(* IEC 61131-3 sources: SortJet_MasterSPS_Aufbau.fbsproj/02_Global Variables, 6 files *)

(* ---- Global_Vars.gvl ---- *)
(* METADATA
{
	"v3Meta": {
		"objectGuid": "27064ae7-2a3c-4a30-8168-a3ab5c131298"
	}
}
*)
{attribute 'allow_unqualified_access'}
NAMESPACE Global_Vars
// Vor StationBasisParameter (Slot 310) initialisieren, dort werden bgFALSE/rgNULL verwendet
{attribute 'global_init_slot' := '295'}
VAR_GLOBAL
//-------------------------------------------------------------------------------------------------
// ALLGEMEINE VARIABLEN
//-------------------------------------------------------------------------------------------------

  // Pointer auf alle Antriebe
  pgAntriebe   : ARRAY[0..65] OF Rexroth_ctrlX_Drive_Eckelmann_MC_V01_02_02;
  bgEtherCatOK : BOOL;

  // Aktivieren \ Deaktivieren des SystemChecks
  bgSystemCheck : ARRAY[cERSTER_AUTOMATIKKREIS..cLETZTER_AUTOMATIKKREIS] OF BOOL := [ cANZAHL_AUTOMATIKKREISE(TRUE) ]; // SystemCheck [AutomatikKreis 1]: FALSE -> Der SystemCheck wird sofort quittiert  TRUE -> SystemCheck wird normal ausgefuehrt

  // Prüfung ob Reset in einem AK aktiv ist
  agbResetAktiv : ARRAY [cERSTER_AUTOMATIKKREIS..cLETZTER_AUTOMATIKKREIS] OF BOOL;

  bgSimulationSiKreisGeschlossen : ARRAY[cERSTER_SICHERHEITSKREIS..cLETZTER_SICHERHEITSKREIS] OF BOOL; // Damit synchronisiert wird, müssen die SKs geschlossen sein - da dies manchmal nicht gegeben ist, kann hiermit

  bgMeldungStromschienenUeberbrueckung : BOOL := FALSE;

  wgStatusPuffer101Oben    : WORD;
  wgStatusPuffer102Unten   : WORD;
  wgStatusPuffer103Oben    : WORD;
  wgStatusPuffer104Unten   : WORD;
  wgStatusTorOben          : WORD;
  wgStatusTorUnten         : WORD;
  // Override für ALLE Achsen - 100 = 100% ; 50 = 50% ;
  rgMaschinenGeschwindigkeitsOverride : REAL := 100;

  (* Hinweis:
     - Pointer- Konstanten [Muessen Global definiert werden]
       => Nicht veraendern
  *)
  bgShuttleEintransportSperren             : ARRAY[cERSTES_SHUTTLE..cLETZTES_SHUTTLE] OF BOOL;
  bgShuttleAustransportSperren             : ARRAY[cERSTES_SHUTTLE..cLETZTES_SHUTTLE] OF BOOL;

  (* Hinweis:
     - Pointer- Konstanten [Muessen Global definiert werden]
       => Nicht veraendern
  *)
  bgTRUE      : BOOL  := TRUE;
  bgFALSE     : BOOL  := FALSE;
  rgNULL      : REAL  := 0;
  wgNULL      : WORD  := 0;

  (* Hinweis:
     - Das Log-Level bestimmt ob und wie die Fehlermeldung geworfen werden->
       Level 0 :=  Nur die übergeordneteten Bausteine werfen einen Fehler
       Level 1 :=  Übergeordnetete Bausteine + Station werfen einen Fehler
       Level 2 :=  Übergeordnetete Bausteine + Station + Unterbausteine werfen einen Fehler
  *)
  wgLogLevel : WORD := 0;
  bgTSLog    : BOOL := TRUE;

  bgStepLogging : BOOL := FALSE;

  Visu_Start_Auto          : BOOL;
  Visu_Notaus_OK           : BOOL := FALSE;

  // Globale Einstellungen
  bgInitialisierungUeberbruecken           : BOOL := FALSE; // Init überspringen
  bgInbetriebnahmeBit                      : BOOL := FALSE; // Inbetriebnahme de/aktivieren
  bgHornAktivieren                         : BOOL := FALSE;  // Horn / Hupe an der Anlage de/aktivieren
  bgSicherheitstechnikBruecken             : BOOL := FALSE; // Inbetriebnahme de/aktivieren
  bgMMIBruecken                            : BOOL := FALSE;
  bgDeaktiviereWatchIOs                    : BOOL := FALSE;
  bgSPS_SIMULATION                         : BOOL := FALSE;
  rgSimScheibenlaenge                      : REAL := 1000.0; // Simulation (bgSPS_SIMULATION): virtuelle Scheibenlaenge [mm] fuer Scheibenmessung und Restwegmessung der simulierten Antriebe
  bgTransfershuttleVortransportAktivieren  : BOOL := FALSE;  // Quittierung des Vortransportauftrags (Ohne Ablauf)
  bgNotHalt_SPS_OK                         : BOOL := TRUE;

  // Ausgaenger - Blink -
  gbFlashbit02sec  : BOOL;
  gbFlashbit05sec  : BOOL;
  gbFlashbit1sec   : BOOL;
  gbFlashbit03sec  : BOOL;
  gbFlashbit12sec  : BOOL;

  // Verfahrueberwachung
  abgVerfahrfreigabeShuttle                    : ARRAY[cERSTES_SHUTTLE..cLETZTES_TRANSFERSHUTTLE] OF BOOL;

  // Init
  M_Init_Ok        : BOOL;

  // Automatikkreise [Speicher - Shuttle - Transfershuttle - ggf. Perepherie
  M_Automatik_Aktiv                         : ARRAY[cERSTER_AUTOMATIKKREIS..cLETZTER_AUTOMATIKKREIS] OF BOOL;
  tonAutomatik_Aktiv                        : ARRAY[cERSTER_AUTOMATIKKREIS..cLETZTER_AUTOMATIKKREIS] OF TON;

  // SystemCheck:
  //   - neue Strukturen aufrufen
  abgDateStationCheck  : ARRAY[101..cLETZTE_STATION, cWAND_1..cANZAHL_WAENDE] OF Auftragsdaten_ST; // Daten die fuer den SystemCheck gebraucht werden

//-------------------------------------------------------------------------------------------------
// ALLGEMEINE STRUKTUREN
//-------------------------------------------------------------------------------------------------
  igIndexFaecherwagenDatenEmpfangen : INT := 0;
  igIndexFaecherwagenDatenSenden    : INT := 0;

  (* Hinweis:
     - Puffer in der Shuttlebahn
  *)
  wgStatusPuffer                       : ARRAY[cERSTES_SHUTTLE..cLETZTES_SHUTTLE] OF WORD;

  (* Hinweis:
     - Allgemeine Konstanten aus der Mathematik
  *)
// *************************************************************************************************
  (* Hinweis:
     - Allgemeine Konstanten aus der Mathematik
  *)
  Mathe : CONSTANTS_MATH;

//-------------------------------------------------------------------------------------------------
// HANDFUNKTIONEN
//-------------------------------------------------------------------------------------------------

  // STATION
  adwgHandfunktionenStationen             : ARRAY[cERSTE_STATION..cLETZTE_STATION] OF DWORD;

  // SHUTTLE
  adwgHandfunktionenShuttle               : ARRAY[cERSTES_SHUTTLE..cLETZTES_SHUTTLE] OF DWORD;

  // TRANSFERSHUTTLE
  adwgHandfunktionenTransfershuttle       : ARRAY[cERSTES_TRANSFERSHUTTLE..cLETZTES_TRANSFERSHUTTLE] OF DWORD;

  // FAECHERWAGENSTATION
  adwgHandfunktionenFaecherwagenStationen : ARRAY[cERSTE_FAECHERWAGENSTATIONS_NR..cLETZTE_FAECHERWAGENSTATIONS_NR] OF DWORD;

//-------------------------------------------------------------------------------------------------
// SYSTEMCHECK
//-------------------------------------------------------------------------------------------------
  wgAnzahlSystemcheckZyklen              : WORD; //  Wird automatisch erkannt

END_VAR
END_NAMESPACE

(* ---- Konstanten.gvl ---- *)
(* METADATA
{
	"v3Meta": {
		"objectGuid": "aefcf88b-f8e6-4fd5-9d29-077a37aead0e"
	}
}
*)
{attribute 'allow_unqualified_access'}
NAMESPACE Konstanten
VAR_GLOBAL CONSTANT

  // Konstanten für die Profibus Master (falls mehrere vorhanden sind)
  cPROFIBUSMASTER_1 : BYTE := 0;
  cPROFIBUSMASTER_2 : BYTE := 1;

  // Konstanten als Ersatz für sizeof
  cSizeOfByte  : WORD := 1;
  cSizeOfWord  : WORD := 2;
  cSizeOfDWord : WORD := 4;
  cSizeOfSInt  : WORD := 1;
  cSizeOfUSInt : WORD := 1;
  cSizeOfInt   : WORD := 2;
  cSizeOfUInt  : WORD := 2;
  cSizeOfDInt  : WORD := 4;
  cSizeOfUDInt : WORD := 4;
  cSizeOfReal  : WORD := 0;

  cMillisecToSec    : WORD  := 1000;
  cMillisecToMinute : WORD  := 60000;

//-------------------------------------------------------------------------------------------------
// SYSTEMCHECK
//-------------------------------------------------------------------------------------------------
  cMAX_ANZAHL_SYSTEMCHECKZYKLEN : WORD := 6;

  // Maximale Anzahl konfigurierbarer Ueberwachungsquellen fuer bpShuttleAnhalten pro Shuttle
  cMAX_SHUTTLE_ANHALTEN_QUELLEN  : WORD := 6;

//-------------------------------------------------------------------------------------------------
// BIT- MASKEN
//-------------------------------------------------------------------------------------------------

  (* Hinweis:
     - Bit Maske
  *)
  // 5432109876543210 ---
  Maske_Bit_0  : WORD := 2#0000000000000001 ;
  Maske_Bit_1  : WORD := 2#0000000000000010 ;
  Maske_Bit_2  : WORD := 2#0000000000000100 ;
  Maske_Bit_3  : WORD := 2#0000000000001000 ;
  Maske_Bit_4  : WORD := 2#0000000000010000 ;
  Maske_Bit_5  : WORD := 2#0000000000100000 ;
  Maske_Bit_6  : WORD := 2#0000000001000000 ;
  Maske_Bit_7  : WORD := 2#0000000010000000 ;
  Maske_Bit_8  : WORD := 2#0000000100000000 ;
  Maske_Bit_9  : WORD := 2#0000001000000000 ;
  Maske_Bit_10 : WORD := 2#0000010000000000 ;
  Maske_Bit_11 : WORD := 2#0000100000000000 ;
  Maske_Bit_12 : WORD := 2#0001000000000000 ;
  Maske_Bit_13 : WORD := 2#0010000000000000 ;
  Maske_Bit_14 : WORD := 2#0100000000000000 ;
  Maske_Bit_15 : WORD := 2#1000000000000000 ;

  // ### KONFIGURIEREN ###

  (* Hinweis:
     - Die folgende Constante darf nicht vergrößert werden, weil es sonst zu einem
       Ueberlauf in der Nachrichtenstruktur kommt
  *)
  cMaxScheibenBeiScheibenMessung  : WORD := 10;

  cMELDUNGScheibe                 : WORD := 0;
  cMAXSCHEIBE                     : WORD := 4;
  cDEFAULTSCHEIBE                 : WORD := 5;
  cMODELLSCHEIBE                  : WORD := 6;

  cGLASDICKEBIS16MM               : WORD := 10;
  cGLASDICKEBIS23MM               : WORD := 11;
  cGLASDICKEBIS29MM               : WORD := 12;

  GLASSTAERKE_DEFAULT_MIN         : WORD := WORD#3;
  GLASSTAERKE_DEFAULT_MAX         : WORD := WORD#14;

  // FAECHERWAGENSTATION
  cEINSCHLEUSESTATION : WORD := 1;
  cPUFFERSTATION      : WORD := 2;
  cFUELLSTATION       : WORD := 3;
  cAUSSCHLEUSESTATION : WORD := 4;
  cKIPPSTATION        : WORD := 5;
  cHUBSTATION         : WORD := 6;
  cENTNAHMESTATION: BOOL := TRUE;

  (* Hinweis:
     - Konstanten fuer das Drehkreuz
  *)
  cGLASDEFAULT : WORD := 0;
  cGLASDREHEN  : WORD := 1;

  (* Hinweis:
     - Grad-Konstanten fuer das Drehkreuz
  *)
  cPOSITION_0Grad    : WORD := 0;
  cPOSITION_90Grad   : WORD := 90;
  cPOSITION_180Grad  : WORD := 180;
  cPOSITION_270Grad  : WORD := 270;
  cPOSITION_360Grad  : WORD := 360;
  rgPOSITION_0Grad   : REAL := REAL#0;
  rgPOSITION_90Grad  : REAL := REAL#90;
  rgPOSITION_180Grad : REAL := REAL#180;
  rgPOSITION_270Grad : REAL := REAL#270;
  rgPOSITION_360Grad : REAL := REAL#360;

  (* Hinweis:
     - Modus wie der FB den Antrieb ansteuern soll
  *)
  cMODUS_MASTER_SLAVE : BYTE := 0;
  cMODUS_HAND         : BYTE := 1;
  cMODUS_RESTWEG      : BYTE := 2;

  (* Hinweis:
     - Unterscheidung Speicher-Einlaufbereich und Speicher-Auslaufbereich
  *)
  cSPEICHER_EINLAUFSEITE : BYTE := 1;
  cSPEICHER_AUSLAUFSEITE : BYTE := 2;

  // Zuweisungskonstanten
  cNULL              : WORD := 0;
  cNULL_WORD_ARRAY   : ARRAY [0..3] OF WORD  :=[ 4(0)];
  cNULL_DWORD_ARRAY  : ARRAY [0..3] OF DWORD :=[ 4(0)];

  cFUEHRUNGSWAGEN    : WORD := 1;
  cZAHNSTANGE        : WORD := 2;

  cSCHMIERKREIS_1    : WORD := 1;
  cSCHMIERKREIS_2    : WORD := 2;
  cSCHMIERKREIS_1_2  : WORD := 3;

//-------------------------------------------------------------------------------------------------
// FOLGEAUFTRAGSTYPEN
//-------------------------------------------------------------------------------------------------
  cFOLGEAUFTRAG_NICHT_AKTIV : WORD := 0;
  cFOLGEAUFTRAG_AKTIV       : WORD := 1;

//-------------------------------------------------------------------------------------------------
// S T A R T - Beladungs- Typ fuer die Shuttle / Stationen nach einem SystemCheck
//-------------------------------------------------------------------------------------------------
  cSTATUS_STATION_FREI              : WORD := 0;
  cSTATUS_STATION_BELEGT            : WORD := 1;
  cSTATUS_STATION_BELEGT_NACHFOLGER : WORD := 2;
  cSTATUS_STATION_BELEGT_VORGEANGER : WORD := 3;

//-------------------------------------------------------------------------------------------------
// BIT-ZUGRIFF WAENDE
//-------------------------------------------------------------------------------------------------
  (* Hinweis:
     - Statuswort <wLetzteScheibe> / <wErsteScheibe>
     - Globale Konstanetn fuer den <bitaccess> der Strukturen ErsteScheibe_ST und LetzteScheibe_ST
     - Werde sind Bit-Codiert
  *)
  cBIT_WAND1   : INT := 0 ;
  cBIT_WAND2   : INT := 1 ;
  cBIT_WAND3   : INT := 2 ;
  cBIT_WAND4   : INT := 3 ;
  cBIT_WAND5   : INT := 4 ;
  cBIT_WAND6   : INT := 5 ;
  cBIT_WAND7   : INT := 6 ;
  cBIT_WAND8   : INT := 7 ;
  cBIT_WAND9   : INT := 8 ;
  cBIT_WAND10  : INT := 9 ;
  cBIT_WAND11  : INT := 10;
  cBIT_WAND12  : INT := 11;
  cBIT_WAND13  : INT := 12;
  cBIT_WAND14  : INT := 13;
  cBIT_WAND15  : INT := 14;
  cBIT_WAND16  : INT := 15;

  (* Hinweis:
     - Bit-Definition für die Auftragsinformationen
  *)
  cBIT_AUFTRAGSTYP          : WORD := 0;
  cBIT_SRCSTATION_EMPTY     : WORD := 1;
  cBIT_Reserve              : WORD := 2;
  cBIT_WALL_1_EMPTY         : WORD := 3;
  cBIT_WALL_2_EMPTY         : WORD := 4;
  cBIT_WALL_3_EMPTY         : WORD := 5;
  cBIT_WALL_4_EMPTY         : WORD := 6;
  cBIT_SRC_WALL_1_EMPTY     : WORD := 7;
  cBIT_SRC_WALL_2_EMPTY     : WORD := 8;
  cBIT_UNUSED               : WORD := 9;
  cBIT_BUFFERSLOT_THICKNESS : WORD := 10;

//-------------------------------------------------------------------------------------------------
// Sensorfehlertypen
//-------------------------------------------------------------------------------------------------

  cAUSNAHMESITUATION_KEIN_SENSOR            : WORD := 0;
  cAUSNAHMESITUATION_EINLAUFSENSOR          : WORD := 1;
  cAUSNAHMESITUATION_AUSLAUFSENSOR          : WORD := 2;
  cAUSNAHMESITUATION_EINLAUF_AUSLAUF_SENSOR : WORD := 3;

//-------------------------------------------------------------------------------------------------
// Status Auftrag
//-------------------------------------------------------------------------------------------------

  cAUFTRAG_FEHLER      : BYTE := 0;
  cAUFTRAG_ERFOLGREICH : BYTE := 1;
  cAUFTRAG_KEIN_STATUS : BYTE := 99;

//-------------------------------------------------------------------------------------------------
// String- Verarbeitung
//-------------------------------------------------------------------------------------------------

   cLINE_FEED       : BYTE := BYTE#16#0A;
   cCARRIAGE_RETURN : BYTE := BYTE#16#0D;

//-------------------------------------------------------------------------------------------------
// ASCII TABELLE
//-------------------------------------------------------------------------------------------------

  (* Hinweis:
     - Datenwoerter in String konvertieren
  *)
  ascii : ARRAY[0..255] OF STRING(1) :=[ 33(' '), '!', '"','#','$$' ,'%' ,'&' ,' ','(' ,')' ,'*' ,'+' ,',' ,
                                        '-' ,'.' ,'/' ,'0' ,'1' ,'2' ,'3' ,'4' ,'5' ,'6' ,'7' ,'8' ,'9' ,':' ,
                                        ';' ,'<' ,'=' ,'>' ,'?' , '@','A' ,'B' ,'C' ,'D' ,'E' ,'F' ,'G' ,'H' ,
                                        'I' ,'J' ,'K' ,'L' ,'M' ,'N' ,'O' ,'P' ,'Q' ,'R' ,'S' ,'T' ,'U' ,'V' ,
                                        'W' ,'X' ,'Y' ,'Z' ,'[','\' ,']' ,'^' ,'_' ,'`' ,'a' ,'b' ,'c' ,'d' ,'e' ,
                                        'f' ,'g' ,'h' ,'i' ,'j' ,'k' ,'l' ,'m' ,'n' ,'o' ,'p' ,'q' ,'r' ,'s' ,'t' ,
                                        'u' ,'v' ,'w' ,'x' ,'y' ,'z' ,'{' ,'|' ,'}' ,'~'];

//-------------------------------------------------------------------------------------------------
// Globale Konstanetn
//-------------------------------------------------------------------------------------------------
  cEVENT_STATUS_STATION_BELADEN         : WORD := 16#1;
  cEVENT_STATUS_FREIGEGEBEN             : WORD := 16#2;
  cEVENT_STATUS_GLAS_NICHT_FREIGEGEBEN  : WORD := 16#4;
  cEVENT_STATUS_QUITTUNG_ISO_LINE_EVENT : WORD := 16#8;
  cEVENT_STATUS_GLASBRUCH               : WORD := 16#10;
  cEVENT_STATUS_GLASABGENOMMEN          : WORD := 16#20;

//-------------------------------------------------------------------------------------------------
// IO am Umrichter
//-------------------------------------------------------------------------------------------------

  // DI an XG31
  cXG31_1_I_1     : WORD  := 16;
  cXG31_2_I_2     : WORD  := 17;
  cXG31_3_I_3     : WORD  := 18;
  cXG31_6_I_4     : WORD  := 19;
  cXG31_7_I_5     : WORD  := 20;
  cXG31_8_I_6_O_1 : WORD  := 21;

  // DI an XG37
  cXG37_1_IO_1    : WORD  := 22;
  cXG37_2_IO_2    : WORD  := 23;

  cXG37_3_I_5     : WORD  := 26;
  cXG37_4_I_6     : WORD  := 27;
  cXG37_5_I_7     : WORD  := 28;
  cXG37_6_I_8     : WORD  := 29;

  // DO an XG37              Die Bits aus dem SignalSteuerwort!
  cXG37_IO_3      : WORD  := 3;
  cXG37_IO_4      : WORD  := 4;
  cXG37_O_5       : WORD  := 5;
  cXG37_O_6       : WORD  := 6;
  cXG37_O_7       : WORD  := 7;
  cXG37_O_8       : WORD  := 8;

END_VAR

END_NAMESPACE

(* ---- MKs.gvl ---- *)
(* METADATA
{
	"v3Meta": {
		"objectGuid": "9b7f8e64-81bc-45e3-b4d2-38b14b6ecc92"
	}
}
*)
{attribute 'allow_unqualified_access'}
NAMESPACE MKs
VAR_GLOBAL
  bgMkParameterOk      : BOOL := FALSE;
END_VAR
END_NAMESPACE

(* ---- PhasenBausteine.gvl ---- *)
(* METADATA
{
	"v3Meta": {
		"objectGuid": "8f2e3603-2a31-4ec8-bbc8-8d5b1492922a"
	}
}
*)
{attribute 'allow_unqualified_access'}
NAMESPACE PhasenBausteine
VAR_GLOBAL CONSTANT

  // UEBERWACHUNG DER SENSORIK
  SENSORIKUEBERWACHUNG_FEHLER                   : INT := -1;
  SENSORIKUEBERWACHUNG_IDLE                     : INT := 0;
  SENSORIKUEBERWACHUNG_INITIALISIERUNG          : INT := 1;
  SENSORIKUEBERWACHUNG_AKTIV                    : INT := 2;
  SENSORIKUEBERWACHUNG_EINLAUFSENSOR_FREIFAHREN : INT := 3;
  SENSORIKUEBERWACHUNG_AUSLAUFSENSOR_FREIFAHREN : INT := 4;
  SENSORIKUEBERWACHUNG_ABGESCHLOSSEN            : INT := 5;

  // TRANSFERSHUTTLE SPEICHERFACH VALIDIERUNG
  SPEICHERFACHVALIDIERUNG_FEHLER                : INT := -1;
  SPEICHERFACHVALIDIERUNG_IDLE                  : INT := 0;
  SPEICHERFACHVALIDIERUNG_INIT                  : INT := 1;
  SPEICHERFACHVALIDIERUNG_AKTIV                 : INT := 2;
  SPEICHERFACHVALIDIERUNG_ABGESCHLOSSEN         : INT := 3;

END_VAR

END_NAMESPACE

(* ---- StationsKonstanten.gvl ---- *)
(* METADATA
{
	"v3Meta": {
		"objectGuid": "160674d4-fa8a-4395-ad23-cbe43462ea3f"
	}
}
*)
{attribute 'allow_unqualified_access'}
NAMESPACE StationsKonstanten
VAR_GLOBAL CONSTANT
 // 5432109876543210
 cStationHandbetrieb : WORD := 2#0000000000000000;
 cStationReset       : WORD := 2#0000000000000001;
 cStationCheck       : WORD := 2#0000000000000010;
 cStationAutomatik   : WORD := 2#0000000000000100;
 cStationReferenz    : WORD := 2#0000000000001000;

 cEinzelStationsCheck       : WORD := 2#0000000000000000;
 cMehrfachStationsCheckTyp1 : WORD := 2#0000000000000001;
 cMehrfachStationsCheckTyp2 : WORD := 2#0000000000000010;
 cMehrfachStationsCheckTyp3 : WORD := 2#0000000000000011;
END_VAR

END_NAMESPACE

(* ---- VISU_VARS.gvl ---- *)
(* METADATA
{
	"v3Meta": {
		"objectGuid": "ca97481c-3185-43db-a213-215d556851fe"
	}
}
*)
{attribute 'allow_unqualified_access'}
NAMESPACE VISU_VARS
VAR_GLOBAL

  wgvisushuttlefehlernr  : WORD;

  bgVisu2StationenDrehrichtungWechsel : BOOL;

  abgVISUFreigabeFremdanlage                 : ARRAY[cERSTE_FREMDANLAGE_AUSLAUF..cLETZTE_FREMDANLAGE_EINLAUF] OF BOOL;

  bgVISUAutomatikModusStation                : ARRAY[cERSTE_STATION..cLETZTE_STATION] OF BOOL;
  bgVISUAutomatikModusShuttle                : ARRAY[cERSTES_SHUTTLE..cLETZTES_TRANSFERSHUTTLE] OF BOOL;

  bgVISUGeblaese                             : ARRAY[cERSTES_SHUTTLE..cLETZTE_STATION, cWAND_1..cANZAHL_WAENDE] OF BOOL;
  bgVISUDrosselklappeAUF                     : ARRAY[cERSTES_SHUTTLE..cLETZTE_STATION] OF BOOL;

  bgVISUGlastransportVor                     : ARRAY[cERSTES_SHUTTLE..cLETZTE_STATION, cWAND_1..cANZAHL_WAENDE] OF BOOL;
  bgVISUGlastransportZurueck                 : ARRAY[cERSTES_SHUTTLE..cLETZTE_STATION, cWAND_1..cANZAHL_WAENDE] OF BOOL;
  bgVISUGlastransportYVor                    : ARRAY[cERSTE_STATION..cLETZTE_STATION] OF BOOL;   // Eckuebergabe: Glastransport Y vor
  bgVISUGlastransportYZurueck                : ARRAY[cERSTE_STATION..cLETZTE_STATION] OF BOOL;   // Eckuebergabe: Glastransport Y zurueck

  // HANDFUNKTIONEN: GREIFER (nur Shuttle, je Wand; Tipptaster der Visu "Handbetrieb Speicher")
  bgVISUGreiferVor                           : ARRAY[cERSTES_SHUTTLE..cLETZTES_SHUTTLE, cWAND_1..cANZAHL_WAENDE] OF BOOL; // Greiferachse vor
  bgVISUGreiferZurueck                       : ARRAY[cERSTES_SHUTTLE..cLETZTES_SHUTTLE, cWAND_1..cANZAHL_WAENDE] OF BOOL; // Greiferachse zurueck
  bgVISUGreiferReferenz                      : ARRAY[cERSTES_SHUTTLE..cLETZTES_SHUTTLE, cWAND_1..cANZAHL_WAENDE] OF BOOL; // Greiferachse referenzieren
  bgVISUGreiferAusfahren                     : ARRAY[cERSTES_SHUTTLE..cLETZTES_SHUTTLE, cWAND_1..cANZAHL_WAENDE] OF BOOL; // Greifer zum Glas ausfahren
  bgVISUGreiferEinfahren                     : ARRAY[cERSTES_SHUTTLE..cLETZTES_SHUTTLE, cWAND_1..cANZAHL_WAENDE] OF BOOL; // Greifer einfahren
  bgVISUGreiferZangeSchliessen               : ARRAY[cERSTES_SHUTTLE..cLETZTES_SHUTTLE, cWAND_1..cANZAHL_WAENDE] OF BOOL; // Greiferzange schliessen
  bgVISUGreiferZangeOeffnen16mm              : ARRAY[cERSTES_SHUTTLE..cLETZTES_SHUTTLE, cWAND_1..cANZAHL_WAENDE] OF BOOL; // Greiferzange oeffnen 16 mm
  bgVISUGreiferZangeOeffnen23mm              : ARRAY[cERSTES_SHUTTLE..cLETZTES_SHUTTLE, cWAND_1..cANZAHL_WAENDE] OF BOOL; // Greiferzange oeffnen 23 mm
  bgVISUGreiferZangeOeffnen29mm              : ARRAY[cERSTES_SHUTTLE..cLETZTES_SHUTTLE, cWAND_1..cANZAHL_WAENDE] OF BOOL; // Greiferzange oeffnen 29 mm
  bgVISUGreiferGlasRueckhalterAusfahren      : ARRAY[cERSTES_SHUTTLE..cLETZTES_SHUTTLE, cWAND_1..cANZAHL_WAENDE] OF BOOL; // Glasrueckhalter (Haltebuegel) ausfahren

  bgVISUQuerfahrtVor                         : ARRAY[cERSTES_SHUTTLE..cLETZTE_STATION] OF BOOL;
  bgVISUQuerfahrtZurueck                     : ARRAY[cERSTES_SHUTTLE..cLETZTE_STATION] OF BOOL;
  bgVISUQuerfahrtReferenz                    : ARRAY[cERSTES_SHUTTLE..cLETZTE_STATION] OF BOOL;
  bgVISUQuerfahrtEintransportPos1            : ARRAY[cERSTES_SHUTTLE..cLETZTE_STATION] OF BOOL;
  bgVISUQuerfahrtAustransportPos1            : ARRAY[cERSTES_SHUTTLE..cLETZTE_STATION] OF BOOL;

  bgVISUVerfahreShuttle                      : ARRAY[cERSTES_SHUTTLE..cLETZTE_STATION] OF BOOL;

  bgVISUAnschlaegeAuf                        : ARRAY[cERSTE_STATION..cLETZTE_STATION] OF BOOL;
  bgVISUAnschlaegeAb                         : ARRAY[cERSTE_STATION..cLETZTE_STATION] OF BOOL;

// Hicham Aenderung vom 25.05.2022: Neue Visu Variablen fuer Handfunktion
  bgVISUHubrahmenAuf_Ebene1                  : ARRAY[cERSTE_STATION..cLETZTE_STATION] OF BOOL;   // Um die zylinder 1 zu steuern: Heben  Ebene 1
  bgVISUHubrahmenAb_Ebene1                   : ARRAY[cERSTE_STATION..cLETZTE_STATION] OF BOOL;   // Um die zylinder 1 zu steuern: Senken Ebene 1
  bgVISUHubrahmenAuf_Ebene2                  : ARRAY[cERSTE_STATION..cLETZTE_STATION] OF BOOL;   // Um die zylinder 2 zu steuern: Heben  Ebene 2
  bgVISUHubrahmenAb_Ebene2                   : ARRAY[cERSTE_STATION..cLETZTE_STATION] OF BOOL;   // Um die zylinder 2 zu steuern: Senken Ebene 2

  bgVISUTransportsperreRunter                : ARRAY[cERSTE_STATION..cLETZTE_STATION] OF BOOL;
  bgVISUTransportsperreHoch                  : ARRAY[cERSTE_STATION..cLETZTE_STATION] OF BOOL;

  bgVISUZentralschmierungStarten             : ARRAY[cERSTES_SHUTTLE..cLETZTES_TRANSFERSHUTTLE] OF BOOL;

  // HANDFUNKTIONEN: HOEHENKONTROLLE
  bgVISUHoehenkontrolleVor                   : ARRAY[cERSTE_STATION..cLETZTE_STATION] OF BOOL;
  bgVISUHoehenkontrolleZurueck               : ARRAY[cERSTE_STATION..cLETZTE_STATION] OF BOOL;
  bgVISUHoehenkontrolleReferenz              : ARRAY[cERSTE_STATION..cLETZTE_STATION] OF BOOL;

  // HANDFUNKTIONEN: DREHEN
  bgVISUDrehen0Grad                          : ARRAY[cERSTE_STATION..cLETZTE_STATION] OF BOOL;
  bgVISUDrehen90Grad                         : ARRAY[cERSTE_STATION..cLETZTE_STATION] OF BOOL;
  bgVISUDrehen180Grad                        : ARRAY[cERSTE_STATION..cLETZTE_STATION] OF BOOL;
  bgVISUDrehen270Grad                        : ARRAY[cERSTE_STATION..cLETZTE_STATION] OF BOOL;
  bgVISUDrehenWechsel                        : ARRAY[cERSTE_STATION..cLETZTE_STATION] OF BOOL;
  bgVISUDrehenReferenz                       : ARRAY[cERSTE_STATION..cLETZTE_STATION] OF BOOL;

  // HANDFUNKTIONEN: KIPPEN
  bgVISUKippen_0_Grad                        : ARRAY[cERSTES_SHUTTLE..cLETZTE_STATION] OF BOOL;
  bgVISUKippen_1_5_Grad                      : ARRAY[cERSTES_SHUTTLE..cLETZTE_STATION] OF BOOL;
  bgVISUKippen_90_Grad                       : ARRAY[cERSTES_SHUTTLE..cLETZTE_STATION] OF BOOL;
  bgVISUKippen_84_Grad                       : ARRAY[cERSTES_SHUTTLE..cLETZTE_STATION] OF BOOL;
  bgVISUKippen_88_5_Grad                     : ARRAY[cERSTES_SHUTTLE..cLETZTE_STATION] OF BOOL;
  bgVISUKippenW1Hoch                         : ARRAY[cERSTES_SHUTTLE..cLETZTE_STATION] OF BOOL;
  bgVISUKippenW1Runter                       : ARRAY[cERSTES_SHUTTLE..cLETZTE_STATION] OF BOOL;
  bgVISUKippenW1Referenz                     : ARRAY[cERSTES_SHUTTLE..cLETZTE_STATION] OF BOOL;
  bgVISUKippenW2Hoch                         : ARRAY[cERSTES_SHUTTLE..cLETZTE_STATION] OF BOOL;
  bgVISUKippenW2Runter                       : ARRAY[cERSTES_SHUTTLE..cLETZTE_STATION] OF BOOL;
  bgVISUKippenW2Referenz                     : ARRAY[cERSTES_SHUTTLE..cLETZTE_STATION] OF BOOL;
  bgVISUKippenW3Hoch                         : ARRAY[cERSTES_SHUTTLE..cLETZTE_STATION] OF BOOL;
  bgVISUKippenW3Runter                       : ARRAY[cERSTES_SHUTTLE..cLETZTE_STATION] OF BOOL;
  bgVISUKippenW3Referenz                     : ARRAY[cERSTES_SHUTTLE..cLETZTE_STATION] OF BOOL;
  bgVISUKippenBremseLoesen                   : ARRAY[cERSTES_SHUTTLE..cLETZTE_STATION] OF BOOL;

  bgVISUKippenGrundstellung                  : ARRAY[cERSTES_SHUTTLE..cLETZTE_STATION] OF BOOL;
  bgVISUKippenUebergabePosition              : ARRAY[cERSTES_SHUTTLE..cLETZTE_STATION] OF BOOL;
  bgVISUKippenReferenz                       : ARRAY[cERSTES_SHUTTLE..cLETZTE_STATION] OF BOOL;

  // HANDFUNKTIONEN: HUB WAND 1
  bgVISUHubW1Auf                             : ARRAY[cERSTE_STATION..cLETZTE_STATION] OF BOOL;
  bgVISUHubW1Ab                              : ARRAY[cERSTE_STATION..cLETZTE_STATION] OF BOOL;
  bgVISUHubW1Referenz                        : ARRAY[cERSTE_STATION..cLETZTE_STATION] OF BOOL;

  bgVISUZylinder1Einfahren                   : ARRAY[cERSTE_STATION..cLETZTE_STATION] OF BOOL;
  bgVISUZylinder2Einfahren                   : ARRAY[cERSTE_STATION..cLETZTE_STATION] OF BOOL;
  bgVISUZylinder1Ausfahren                   : ARRAY[cERSTE_STATION..cLETZTE_STATION] OF BOOL;
  bgVISUZylinder2Ausfahren                   : ARRAY[cERSTE_STATION..cLETZTE_STATION] OF BOOL;

  // HANDFUNKTIONEN: HUB ALLGEMEIN
  bgVISUHubPositionW1                        : ARRAY[cERSTE_STATION..cLETZTE_STATION] OF BOOL;
  bgVISUHubPositionW2                        : ARRAY[cERSTE_STATION..cLETZTE_STATION] OF BOOL;
  bgVISUHubPositionNachfolger                : ARRAY[cERSTE_STATION..cLETZTE_STATION] OF BOOL;
  bgVISUHubPositionVorgaenger                : ARRAY[cERSTE_STATION..cLETZTE_STATION] OF BOOL;

  bgVISUGlastransportOeffnungGeschlossen     : ARRAY[cERSTES_SHUTTLE..cLETZTE_STATION, cWAND_1..cANZAHL_WAENDE] OF BOOL;
  bgVISUGlastransportOeffnungMinimal         : ARRAY[cERSTES_SHUTTLE..cLETZTE_STATION, cWAND_1..cANZAHL_WAENDE] OF BOOL;
  bgVISUGlastransportOeffnungMittel          : ARRAY[cERSTES_SHUTTLE..cLETZTE_STATION, cWAND_1..cANZAHL_WAENDE] OF BOOL;
  bgVISUGlastransportOeffnungMaximal         : ARRAY[cERSTES_SHUTTLE..cLETZTE_STATION, cWAND_1..cANZAHL_WAENDE] OF BOOL;

  bgVISUW1QuerverstellungMinimal             : ARRAY[cERSTES_SHUTTLE..cLETZTE_STATION] OF BOOL;
  bgVISUW1QuerverstellungMittel              : ARRAY[cERSTES_SHUTTLE..cLETZTE_STATION] OF BOOL;
  bgVISUW1QuerverstellungMaximal             : ARRAY[cERSTES_SHUTTLE..cLETZTE_STATION] OF BOOL;

  bgVISUSicherungsbolzenEinfahren            : ARRAY[cERSTE_STATION..cLETZTE_STATION] OF BOOL;

  bgVISUZentrierbolzenEinfahren              : ARRAY[cERSTES_SHUTTLE..cLETZTE_STATION] OF BOOL;
  bgVISUZentrierbolzenAusfahren              : ARRAY[cERSTES_SHUTTLE..cLETZTE_STATION] OF BOOL;

  // Transfershuttle (TFS)
  wgVISUAuswahlTransferShuttle               : WORD := 151;
  bgVisuTFSRiemenAnheben                     : ARRAY[cERSTES_TRANSFERSHUTTLE..cLETZTES_TRANSFERSHUTTLE] OF BOOL;
  bgVisuTFSRiemenSenken                      : ARRAY[cERSTES_TRANSFERSHUTTLE..cLETZTES_TRANSFERSHUTTLE] OF BOOL;
  bgVisuTFSAbfrageEinlaufAuf                 : ARRAY[cERSTES_TRANSFERSHUTTLE..cLETZTES_TRANSFERSHUTTLE] OF BOOL;
  bgVisuTFSAbfrageAuslaufAuf                 : ARRAY[cERSTES_TRANSFERSHUTTLE..cLETZTES_TRANSFERSHUTTLE] OF BOOL;
  bgVisuTFSAbfrageEinlaufEin                 : ARRAY[cERSTES_TRANSFERSHUTTLE..cLETZTES_TRANSFERSHUTTLE] OF BOOL;
  bgVisuTFSAbfrageAuslaufEin                 : ARRAY[cERSTES_TRANSFERSHUTTLE..cLETZTES_TRANSFERSHUTTLE] OF BOOL;
  bgVisuTFS_BreiteAbfrageEinlaufAuf          : ARRAY[cERSTES_TRANSFERSHUTTLE..cLETZTES_TRANSFERSHUTTLE] OF BOOL;
  bgVisuTFS_BreiteAbfrageAuslaufAuf          : ARRAY[cERSTES_TRANSFERSHUTTLE..cLETZTES_TRANSFERSHUTTLE] OF BOOL;
  bgVisuTFS_BreiteAbfrageEinlaufEin          : ARRAY[cERSTES_TRANSFERSHUTTLE..cLETZTES_TRANSFERSHUTTLE] OF BOOL;
  bgVisuTFS_BreiteAbfrageAuslaufEin          : ARRAY[cERSTES_TRANSFERSHUTTLE..cLETZTES_TRANSFERSHUTTLE] OF BOOL;
  bgVisuTFSScheibeZurueckHolen               : ARRAY[cERSTES_TRANSFERSHUTTLE..cLETZTES_TRANSFERSHUTTLE] OF BOOL;
  bgVisuTFSGlastransporttestAktivieren       : ARRAY[cERSTES_TRANSFERSHUTTLE..cLETZTES_TRANSFERSHUTTLE] OF BOOL;
  bgVisuTFSQuerfahrtVor                      : ARRAY[cERSTES_TRANSFERSHUTTLE..cLETZTES_TRANSFERSHUTTLE] OF BOOL;
  bgVisuTFSQuerfahrtZurueck                  : ARRAY[cERSTES_TRANSFERSHUTTLE..cLETZTES_TRANSFERSHUTTLE] OF BOOL;
  bgVisuTFSQuerfahrtReferenz                 : ARRAY[cERSTES_TRANSFERSHUTTLE..cLETZTES_TRANSFERSHUTTLE] OF BOOL;
  bgVisuTFSZentralschmierungStarten          : ARRAY[cERSTES_TRANSFERSHUTTLE..cLETZTES_TRANSFERSHUTTLE] OF BOOL;

  // HANDFUNKTIONEN: FAECHERWAGEN
  bgVISUFWEntriegelungEinfahren              : ARRAY[cERSTE_FAECHERWAGENSTATIONS_NR..cLETZTE_FAECHERWAGENSTATIONS_NR] OF BOOL;
  bgVISUFWEntriegelungAusfahren              : ARRAY[cERSTE_FAECHERWAGENSTATIONS_NR..cLETZTE_FAECHERWAGENSTATIONS_NR] OF BOOL;
  bgVISUFWGreiferEinfahren                   : ARRAY[cERSTE_FAECHERWAGENSTATIONS_NR..cLETZTE_FAECHERWAGENSTATIONS_NR] OF BOOL;
  bgVISUFWGreiferAusfahren                   : ARRAY[cERSTE_FAECHERWAGENSTATIONS_NR..cLETZTE_FAECHERWAGENSTATIONS_NR] OF BOOL;
  bgVISUFWGegenhalterEinfahren               : ARRAY[cERSTE_FAECHERWAGENSTATIONS_NR..cLETZTE_FAECHERWAGENSTATIONS_NR] OF BOOL;
  bgVISUFWGegenhalterAusfahren               : ARRAY[cERSTE_FAECHERWAGENSTATIONS_NR..cLETZTE_FAECHERWAGENSTATIONS_NR] OF BOOL;
  bgVISUFWLinearEinheitVor                   : ARRAY[cERSTE_FAECHERWAGENSTATIONS_NR..cLETZTE_FAECHERWAGENSTATIONS_NR] OF BOOL;
  bgVISUFWLinearEinheitZurueck               : ARRAY[cERSTE_FAECHERWAGENSTATIONS_NR..cLETZTE_FAECHERWAGENSTATIONS_NR] OF BOOL;
  bgVISUFWLinearEinheitShuttle               : ARRAY[cERSTE_FAECHERWAGENSTATIONS_NR..cLETZTE_FAECHERWAGENSTATIONS_NR] OF BOOL;
  bgVISUFWRolltorHoch                        : ARRAY[cERSTE_FAECHERWAGENSTATIONS_NR..cLETZTE_FAECHERWAGENSTATIONS_NR] OF BOOL;
  bgVISUFWRolltorRunter                      : ARRAY[cERSTE_FAECHERWAGENSTATIONS_NR..cLETZTE_FAECHERWAGENSTATIONS_NR] OF BOOL;
  bgVISUFWQuittierungLichtschranke           : ARRAY[cERSTE_FAECHERWAGENSTATIONS_NR..cLETZTE_FAECHERWAGENSTATIONS_NR] OF BOOL;

  // STATUS: FAECHERWAGEN (alle Varianten; die Visu liest den Status hier statt aus den IOs der Station)
  astgFaecherwagenstatusVisu                 : ARRAY[cERSTE_FAECHERWAGENSTATIONS_NR..cLETZTE_FAECHERWAGENSTATIONS_NR] OF Faecherwagenstatus_Visu_ST;

  bgVISUSetWatchIO                           : BOOL;
  wgVISUWatchIONr                            : WORD;
  bgVISUWatchIOAktiv                         : BOOL;

  bgVisuStart                                : BOOL := FALSE;

  bgVISUFehlerAusloesen                      : BOOL;

  bgVisu2StationenVor                 : BOOL := FALSE;
  bgVisu2StationenZurueck             : BOOL := FALSE;
  iGewaehlteStation1                  : WORD := 101;
  iGewaehlteStation2                  : WORD := 101;
  bgStation1W1                        : BOOL := FALSE;
  bgStation1W2                        : BOOL := FALSE;
  bgStation2W1                        : BOOL := FALSE;
  bgStation2W2                        : BOOL := FALSE;
  bgVISU_EINLAUFSENSOR_STATION_1      : BOOL;
  bgVISU_AUSLAUFSENSOR_STATION_1      : BOOL;
  bgVISU_EINLAUFSENSOR_STATION_2      : BOOL;
  bgVISU_AUSLAUFSENSOR_STATION_2      : BOOL;

  // Antriebsraddurchmesser berechenen

  biDurchmesserIst                    : REAL := 0;
  biDurchmesserSoll                   : REAL := 0;
  biWegIst                            : REAL := 0;
  biWegSoll                           : REAL := 0;
  bgBerechnen                         : BOOL;

  abgStationsstatusVisu               : ARRAY[101..cLETZTE_STATION] OF Stationsstatus_Visu_ST;

// Antriebe verfahren
  bgVisuAntriebeVerfahrenAktiv        : BOOL;
  wgAuswahlAchsID                     : WORD := 0;
  rgZielPos                           : REAL := 0;
  rgGeschwindigkeit                   : REAL := 0;
  wgMasterNummer                      : WORD := 0;

  // Test ofne Einlauflinie
  bgVisuQuittEintransport             : ARRAY [101..cLETZTE_STATION] OF BOOL;

END_VAR

END_NAMESPACE
